(* IEC 61131-3 sources: POMIRTS_lab3/AS/Library_2/AsBrMath, 3 files *)

(* ---- AsBrMath.typ ---- *)
TYPE

END_TYPE

(* ---- AsBrMath.fun ---- *)
{REDUND_OK} FUNCTION brmatan2 : REAL               (*calculates the arc tangent of y/x*)
	VAR_INPUT
		y	:REAL;                     (*y*)
		x	:REAL;                     (*x*)
	END_VAR
END_FUNCTION

{REDUND_OK} FUNCTION brmceil : REAL                (*calculates the smallest integer value which is greater than or equal to the input value*)
	VAR_INPUT
		x	:REAL;                     (*input value*)
	END_VAR
END_FUNCTION

{REDUND_OK} FUNCTION brmcosh : REAL                (*calculates the hyperbolic cosine of x*)
	VAR_INPUT
		x	:REAL;                     (*input value*)
	END_VAR
END_FUNCTION

{REDUND_OK} FUNCTION brmfloor : REAL               (*calculates the largest integer value which is less than or equal to the input value*)
	VAR_INPUT
		x	:REAL;                     (*input value*)
	END_VAR
END_FUNCTION

{REDUND_OK} FUNCTION brmfmod : REAL                (*calculates the remainder of the division x/y*)
	VAR_INPUT
		x	:REAL;                     (*numerator*)
		y	:REAL;                     (*denominator*)
	END_VAR
END_FUNCTION

{REDUND_OK} FUNCTION brmfrexp : REAL               (*calculates the mantissa and the exponent of a floating point number*)
	VAR_INPUT
		x	:REAL;                     (*input value*)
		pExp	:UDINT;                (*address of the exponent (address of DINT) (base 2)*)
	END_VAR
END_FUNCTION

{REDUND_OK} FUNCTION brmldexp : REAL               (*calculates a floating point number from mantissa x and exponent exp*)
	VAR_INPUT
		x	:REAL;                     (*mantissa*)
		exp_val	:DINT;                 (*exponent (base 2)*)
	END_VAR
END_FUNCTION

{REDUND_OK} FUNCTION brmmodf : REAL                (*separates a floating point number into an integer and decimal part*)
	VAR_INPUT
		x	:REAL;                     (*input value*)
		plp	:UDINT;                    (*address of the integer part (address of a REAL value)*)
	END_VAR
END_FUNCTION

{REDUND_OK} FUNCTION brmpow : REAL                 (*calculates x raised to the power of y*)
	VAR_INPUT
		x	:REAL;                     (*base*)
		y	:REAL;                     (*exponent*)
	END_VAR
END_FUNCTION

{REDUND_OK} FUNCTION brmsinh : REAL                (*calculates the hyperbolic sine of x*)
	VAR_INPUT
		x	:REAL;                     (*input value*)
	END_VAR
END_FUNCTION

{REDUND_OK} FUNCTION brmtanh : REAL                (*calculates the hyperbolic tangent of x*)
	VAR_INPUT
		x	:REAL;                     (*input value*)
	END_VAR
END_FUNCTION

(* ---- AsBrMath.var ---- *)
VAR CONSTANT
	brm2_SQRTPI	: REAL	:= 1.12838;        (*2/(square root from PI)*)
	brmSQRT1_2	: REAL	:= 0.707107;       (*square root from 1/2*)
	brmSQRTPI	: REAL	:= 1.77245;        (*square root from PI*)
	brmLOG2_E	: REAL	:= 0.693147;       (*log with the base 2 from E*)
	brmLOG10E	: REAL	:= 0.434294;       (*log with the base 10 from E*)
	brmIVLN10	: REAL	:= 0.434294;       (*1/(ln from 10)*)
	brmINVLN2	: REAL	:=  1.4427;        (*1/(ln from 2)*)
	brmTWOPI	: REAL	:= 6.28319;        (*2 PI*)
	brmSQRT3	: REAL	:= 1.73205;        (*square root from 3*)
	brmSQRT2	: REAL	:= 1.41421;        (*square root from 2*)
	brmLOG2E	: REAL	:=  1.4427;        (*log with the base 2 from E*)
	brmLN2LO	: REAL	:= 1.90821e-010;   (*log with the base 2 from LOW*)
	brmLN2HI	: REAL	:= 0.693147;       (*log with the base 2 from HIGH*)
	brm3PI_4	: REAL	:= 2.35619;        (*3/4 PI*)
	brmPI_4	: REAL	:= 0.785398;           (*PI/4*)
	brmPI_2	: REAL	:=  1.5708;            (*PI/2*)
	brmLN10	: REAL	:= 2.30259;            (*ln from 10*)
	brm2_PI	: REAL	:= 0.63662;            (*2/PI*)
	brm1_PI	: REAL	:= 0.31831;            (*1/PI*)
	brmLN2	: REAL	:= 0.693147;           (*ln from 2*)
	brmPI	: REAL	:= 3.14159;            (*PI*)
	brmE	: REAL	:= 2.71828;            (*E*)
END_VAR
